Fanuc KAREL source: KT00278.KL

PROGRAM KT00278
%NOLOCKGROUP
VAR
  P1: POSITION
  P2: JOINTPOS
  OUT: BOOLEAN
BEGIN
  OUT = P1 = P2
END KT00278
